Staubli VAL3: changeDataLib.pgx

public program changeDataLib(num x_nLib (dimensions=1))
  local num l_nResult
begin
  //形参：x_nLib
  //对应实参：savedata:nLibIndex
  bTosave=true
  call trajectory:onSave(bTosave)
  bTosave=true
  call prog:onSave(bTosave)
  call trajectory:loadTRAJ(x_nLib,l_nResult)
  call prog:loadPROG(x_nLib,l_nResult)

end
